// TIA Portal V20 export
// export: Created 2026-10-12T04:58:22.3823783Z, ExportSetting WithDefaults, DisplayName Totally Integrated Automation Portal, DisplayVersion V20, DisplayName TIA Portal Openness, DisplayVersion V20, DisplayName TIA Portal Teamcenter Gateway, DisplayVersion V20, DisplayName TIA Portal Version Control Interface, DisplayVersion V20, DisplayName SINAMICS Startdrive Advanced, DisplayVersion V20 SP1 Update 2, DisplayName SINAMICS Startdrive G110M, G120, G120C, G120D, G120P, G115D, DisplayVersion V20 SP1 Update 2, DisplayName SINAMICS Startdrive G130, G150, S120, S150, SINAMICS MV, G220, S200, S210, DisplayVersion V20 SP1 Update 2, DisplayName STEP 7 Professional, DisplayVersion V20, DisplayName STEP 7 Safety, DisplayVersion V20, DisplayName WinCC Basic/Comfort/Advanced, DisplayVersion V20, DisplayName WinCC Professional, DisplayVersion V20, DisplayName WinCC Unified, DisplayVersion V20
DATA_BLOCK "GDB_StateAlarmTest"   // DB20
{ S7_Optimized_Access := 'TRUE' }
VERSION : 0.1
// stored: AutoNumber true, DBAccessibleFromOPCUA true, DBAccessibleFromWebserver true, IsOnlyStoredInLoadMemory false, IsRetainMemResEnabled false, IsWriteProtectedInAS false, MemoryReserve 100
   VAR
      ClearLog : Bool;
      RaisePulse : Bool;
      GonePulse : Bool;
      FillPulse : Bool;
      CauseLive : Bool;
      PublishState : Bool;
      StateValue : Bool;
      Position : DInt;
      StateIndex : Int;
      ResetClass : DInt;
      FillCount : Int;
      Diag { S7_SetPoint := 'True'} : "ST_Diagnostic";
      Slot { ExternalWritable := 'False'} : Int;
      GoneAccepted { ExternalWritable := 'False'} : Bool;
      SinkCome { ExternalWritable := 'False'} : UDInt;
      SinkClose { ExternalWritable := 'False'} : UDInt;
      SinkLast { ExternalWritable := 'False'; S7_SetPoint := 'True'} : "ST_AlarmEvent";
      NativeFaultSlot { ExternalWritable := 'False'} : Int;
      StandaloneCount { ExternalWritable := 'False'} : Int;
      StandaloneReturn { ExternalWritable := 'False'} : Bool;
      StandaloneFlags { ExternalWritable := 'False'; S7_SetPoint := 'True'} : Array[1..12] of "ST_StateFlag";
      CauseSlot { ExternalAccessible := 'False'; ExternalVisible := 'False'; ExternalWritable := 'False'} : Int;
      Touched { ExternalAccessible := 'False'; ExternalVisible := 'False'; ExternalWritable := 'False'} : Array[1..12] of Bool;
   END_VAR
BEGIN
END_DATA_BLOCK
